Fanuc KAREL source: kf00103.KL

-- PROVISIONAL review KL for V1013-1; original PC SHA256 ebd53a01a1a195094d654d2b60efd9bcd58a41a82f1ef39e2b11e6c2d3b4cb66
-- Incomplete behavior may be omitted. Consult companion uncertainty JSON. Do not deploy.
PROGRAM KF00103
%NOLOCKGROUP
BEGIN
  -- UNRESOLVED_PC offsets 5-16; opcodes 2E,23
  -- UNRESOLVED_PC offsets 21-32; opcodes 2E,23
  -- UNRESOLVED_PC offsets 37-57; opcodes 27,27,9D,22,2A,22,31
  -- UNRESOLVED_PC offsets 62-66; opcodes 7F
END KF00103
